(* IEC 61131-3 sources: ecmc_plugin_strucpp/examples/psi_ioc_examples/ioc_project_minimal/src/generated, 1 file *)

(* ---- main_bundle.st ---- *)
(* Auto-generated by strucpp_bundle_st.py. *)

(* BEGIN main.st *)
PROGRAM MAIN
VAR
  actual_position    AT %IW0 : INT;   // @ecmc ec.s14.positionActual01
  drive_control      AT %QW0 : WORD;  // @ecmc ec.s14.driveControl01
  velocity_setpoint  AT %QW2 : INT;   // @ecmc ec.s14.velocitySetpoint01
  cycle_counter      AT %MW0 : INT;   // @epics rec=Main-CycleCounterAct
  actual_pos_export          : INT;   // @epics prefix=$(IOC): rec=Main-PosActMini
END_VAR

actual_pos_export := actual_position;
cycle_counter := cycle_counter + 1;
drive_control := 16#0001;

IF actual_position < 0 THEN
  velocity_setpoint := 1000;
ELSIF actual_position > 1000 THEN
  velocity_setpoint := -1000;
END_IF;
END_PROGRAM
(* END main.st *)
